Fanuc KAREL source: KD00022.KL

PROGRAM KD00022
%NOLOCKGROUP
VAR
  I: INTEGER
  J: INTEGER
  B: BOOLEAN
  R: REAL
  S: STRING[80]
  SAVED IN CMOS: INTEGER
BEGIN
  I = 1
END KD00022
